// TIA Portal V21 export
// export: Created 2026-11-08T21:35:35.212555Z, ExportSetting WithDefaults, DisplayName Totally Integrated Automation Portal, DisplayVersion V21 Update 3, DisplayName STEP 7 Professional, DisplayVersion V21 Update 3, DisplayName STEP 7 Safety, DisplayVersion V21, DisplayName Tech WebApplication, DisplayVersion V21, DisplayName WinCC Basic/Comfort/Advanced, DisplayVersion V21 Update 3, DisplayName WinCC Unified, DisplayVersion V21 Update 3
FUNCTION_BLOCK "FB_StlC_040"   // FB93, STL
TITLE = STL call WriteToArrayDBL
{ S7_Optimized_Access := 'TRUE' }
VERSION : 0.1
// stored: AutoNumber true, IsRetainMemResEnabled false, MemoryReserve 100, UDAEnableTagReadback false
   VAR_INPUT
      req : Bool;
      di1 : DInt;
      dba : DB_ANY;
   END_VAR
   VAR_OUTPUT
      busy : Bool;
      done : Bool;
      err : Int;
   END_VAR
   VAR
      val : Int;
      inst { S7_SetPoint := 'True'} : WriteToArrayDBL;
   END_VAR
BEGIN

NETWORK
TITLE = 040 WriteToArrayDBL
      CALL  #inst
      ( req   := #req,
        db    := #dba,
        index := #di1,
        value := #val,
        busy  := #busy,
        done  := #done,
        error := #err
      );
END_FUNCTION_BLOCK
